Staubli VAL3: physicalIO.pgx

program physicalIO()
// Lab2A Level 3 - shared manual simulation / physical cycle
begin

  while true

    // Read sensors.
    partOnTool  = (io:bIn0 == true)
    partAtClass = (io:bIn1 == true)
    partIsMetal = (io:bIn2 == true)
    partAtRamp  = (io:bIn4 == true)

    // Apply output commands; the barrier uses inverted logic.
    io:bOut0 = vacuumOn
    io:bOut1 = blowOn

    io:bOut2 = trolleyOn
    io:bOut3 = nonMetalGate
    io:bOut4 = metalGate
    io:bOut5 = !barrierClosed

    ioReady = true
    delay(0.01)

  endWhile
end
